FUNCTION CheckBounds : DINT
VAR_INPUT
	index, lower, upper : DINT;
END_VAR
VAR
END_VAR

IF index<lower THEN
	CheckBounds := lower;
	Errors:=Errors+1;
ELSIF index>upper THEN
	CheckBounds := upper;
	Errors:=Errors+1;
ELSE
	CheckBounds := index;
END_IF

END_FUNCTION

(* stored: Version 1.1.0.1, ProductVersion 3.1.4024.13
   POU CheckBounds: Id {7f76f90f-81d7-45fd-8a29-3301632c9cab}, SpecialFunc CheckBounds *)
